FUNCTION_BLOCK fb_Dev_AnalogSensor_CurrentTransducer EXTENDS fb_Dev_AnalogSensor
VAR_INPUT
END_VAR
VAR_OUTPUT
END_VAR
VAR
	_cfgShuntResValue	:LREAL;
	_cfgWindingRatio	:LREAL;
END_VAR

DeviceLogic();

scaleInput();

FaultHandler();

setHMI();

stsSensorRawSignal	:= _sensorRawSignal;
stsEngValue			:= _engValue;

PROPERTY cfgShuntResValue : LREAL
GET
cfgShuntResValue := _cfgShuntResValue;
END_GET
SET
_cfgShuntResValue := cfgShuntResValue;
END_SET
END_PROPERTY

PROPERTY cfgWindingRatio : LREAL
GET
cfgWindingRatio := _cfgWindingRatio;
END_GET
SET
_cfgWindingRatio := cfgWindingRatio;
END_SET
END_PROPERTY

(*FB_Init is always available implicitly and it is used primarily for initialization.
The return value is not evaluated. For a specific influence, you can also declare the
methods explicitly and provide additional code there with the standard initialization
code. You can evaluate the return value.*)
METHOD FB_Init : BOOL
VAR_INPUT
	(* TRUE: the retain variables are initialized (reset warm / reset cold)*)
	bInitRetains	: BOOL;
	(* TRUE: the instance will be copied to the copy code afterward (online change)   *)
	bInCopyCode	: BOOL;
	cfgDeviceName		: STRING;
	cfgEnable			: BOOL;
	cfgInitEventClass	: BOOL;
	cfgAlarmEnable		: BOOL;
	cfgAlarmH			: LREAL;
	cfgAlarmHH			: LREAL;
	cfgAlarmL			: LREAL;
	cfgAlarmLL			: LREAL;
	cfgEngUnit			: STRING;
	cfgCalOffset		: LREAL;
	cfgCalGain			: LREAL := 1.0;	// omitted in the declaration = 1 (no correction)
	cfgShuntResValue	: LREAL;
	cfgWindingRatio		: LREAL;
END_VAR
THIS^.cfgDeviceName 		:= 		cfgDeviceName; 		
THIS^.cfgEnable 			:= 	    cfgEnable; 	
THIS^.cfgInitEventClass		:= 		cfgInitEventClass;
THIS^.cfgAlarmEnable		:=		cfgAlarmEnable;
THIS^.cfgAlarmH				:=		cfgAlarmH;
THIS^.cfgAlarmHH			:=		cfgAlarmHH;
THIS^.cfgAlarmL				:=		cfgAlarmL;
THIS^.cfgAlarmLL			:=		cfgAlarmLL;
THIS^.cfgCalOffset			:=		cfgCalOffset;
THIS^.cfgCalGain			:=		cfgCalGain;
THIS^.cfgEngUnit			:=		cfgEngUnit;
THIS^.cfgShuntResValue		:=		cfgShuntResValue;
THIS^.cfgWindingRatio		:=		cfgWindingRatio;

THIS^.HMI.cfgAlarmEnable	:= cfgAlarmEnable;
THIS^.HMI.cfgAlarmH			:= cfgAlarmH;
THIS^.HMI.cfgAlarmHH		:= cfgAlarmHH;
THIS^.HMI.cfgAlarmL			:= cfgAlarmL;
THIS^.HMI.cfgAlarmLL		:= cfgAlarmLL;
THIS^.HMI.cfgEngUnit		:= cfgEngUnit;
THIS^.HMI.cfgCalOffset		:= cfgCalOffset;
THIS^.HMI.cfgCalGain		:= cfgCalGain;
END_METHOD

METHOD scaleInput : BOOL
IF cfgScalingNeeded THEN
	_sensorRawSignal	:= F_AnalogToEngUnit(inpRawIOChannel, cfgChannelMinInt, cfgChannelMaxInt, cfgSensorMin, cfgSensorMax);
	_engValue			:= (_sensorRawSignal * _cfgWindingRatio / _cfgShuntResValue) * _CalGain + _calOffset;
ELSE
	_sensorRawSignal := inpRawIOChannel;
	_engValue		 := (inpRawIOChannel * _CalGain) + _calOffset;
END_IF
END_METHOD

END_FUNCTION_BLOCK

(* stored: Version 1.1.0.1
   POU fb_Dev_AnalogSensor_CurrentTransducer: Id {a822f842-1ccd-4194-bd47-dd8572ada53a}, SpecialFunc None
   Property cfgShuntResValue: Id {6b70de73-49bf-4869-88ef-248a795fb48a}
   Get Get: Id {d311cfd9-361d-4444-ab8a-492a0ed0d0aa}
   Set Set: Id {08985d1b-3f4b-4259-9d83-855bf7d26360}
   Property cfgWindingRatio: Id {b7763c4b-b735-47d4-bd66-ff8104a08d23}
   Get Get: Id {497d4c6d-88d7-4aec-a7cd-23642fa1a4ba}
   Set Set: Id {eca31712-efbd-492a-a4a5-b57d836ff1b7}
   Method FB_Init: Id {4e76c754-8e8c-4f3a-abda-377adc0a0941}
   Method scaleInput: Id {0676921f-fb3f-4c05-a1a0-4a7a7f1ff178} *)
